// TIA Portal V20 export
// export: Created 2026-10-20T18:54:58.074688Z, ExportSetting None, DisplayName Totally Integrated Automation Portal, DisplayVersion V20 Update 6, DisplayName TIA Portal Openness, DisplayVersion V20 Update 6, DisplayName TIA Portal Version Control Interface, DisplayVersion V20 Update 6, DisplayName SINAMICS Startdrive Advanced, DisplayVersion V20 SP1, DisplayName SINAMICS Startdrive G130, G150, S120, S150, SINAMICS MV, G220, S200, S210, DisplayVersion V20 SP1, DisplayName SINAMICS Startdrive G110M, G120, G120C, G120D, G120P, G115D, DisplayVersion V20 SP1, DisplayName STEP 7 Professional, DisplayVersion V20 Update 6, DisplayName STEP 7 Safety, DisplayVersion V20 Update 2, DisplayName WinCC Basic/Comfort/Advanced, DisplayVersion V20 Update 6, DisplayName WinCC Unified, DisplayVersion V20 Update 6
VAR_GLOBAL   // PLC tag table "IO_ET200_2"
   "C2205 - SENSOR CNV RIGHT (PALLET DETECT 1)" AT %I354.4 : Bool;
   "C2204 - SENSOR CNV RIGHT (PALLET DETECT 1)" AT %I352.4 : Bool;
   "C2206 - SENSOR CNV RIGHT (PALLET DETECT 1)" AT %I356.4 : Bool;
   "C2203 - SENSOR CNV RIGHT (PALLET DETECT 1)" AT %I350.4 : Bool;
   "C2208 - SENSOR CNV RIGHT (PALLET DETECT 1)" AT %I360.4 : Bool;
   "KEY REMOTE/LOCAL L7 - CH2(2)" AT %I1654.5 : Bool;
   "E-STOP L7 - CH2(2)" AT %I1654.4 : Bool;
   "KEY REMOTE/LOCAL L8 - CH1(2)" AT %I1654.3 : Bool;
   "KEY REMOTE/LOCAL L6 - CH1(2)" AT %I1646.3 : Bool;
   "KEY REMOTE/LOCAL L7 - CH1(2)" AT %I1654.1 : Bool;
   "KEY REMOTE/LOCAL L2 - CH2(2)" AT %I1476.7 : Bool;
   "E-STOP L3 - CH1(2)" AT %I1638.0 : Bool;
   "KEY REMOTE/LOCAL L3 - CH1(2)" AT %I1638.1 : Bool;
   "E-STOP L4 - CH1(2)" AT %I1638.2 : Bool;
   "KEY REMOTE/LOCAL L4 - CH1(2)" AT %I1638.3 : Bool;
   "E-STOP L3 - CH2(2)" AT %I1638.4 : Bool;
   "KEY REMOTE/LOCAL L3 - CH2(2)" AT %I1638.5 : Bool;
   "E-STOP L4 - CH2(2)" AT %I1638.6 : Bool;
   "KEY REMOTE/LOCAL L4 - CH2(2)" AT %I1638.7 : Bool;
   "E-STOP L5 - CH1(2)" AT %I1646.0 : Bool;
   "KEY REMOTE/LOCAL L5 - CH1(2)" AT %I1646.1 : Bool;
   "E-STOP L6 - CH1(2)" AT %I1646.2 : Bool;
   "E-STOP L5 - CH2(2)" AT %I1646.4 : Bool;
   "KEY REMOTE/LOCAL L5 - CH2(2)" AT %I1646.5 : Bool;
   "E-STOP L6 - CH2(2)" AT %I1646.6 : Bool;
   "KEY REMOTE/LOCAL L6 - CH2(2)" AT %I1646.7 : Bool;
   "E-STOP L7 - CH1(2)" AT %I1654.0 : Bool;
   "E-STOP L8 - CH1(2)" AT %I1654.2 : Bool;
   "E-STOP L2 - CH2(2)" AT %I1476.6 : Bool;
   "KEY REMOTE/LOCAL L2 - CH1(2)" AT %I1476.3 : Bool;
   "E-STOP L2 - CH1(2)" AT %I1476.2 : Bool;
   "E-STOP L8 - CH2(2)" AT %I1654.6 : Bool;
   "KEY REMOTE/LOCAL L8 - CH2(2)" AT %I1654.7 : Bool;
   "C2102 - SENSOR SAFETY PIN1 DOWN" AT %I175.3 : Bool;
   "C2202 - SENSOR CNV LEFT (PALLET DETECT 2)" AT %I270.0 : Bool;
   "CVTD2 SENSOR CONVEYOR CENTER" AT %I1275.5 : Bool;
   "C2206 - SHUTTLE IN POSITION 2" AT %I357.6 : Bool;
   "C2205 - SENSOR SAFETY PIN1 DOWN" AT %I355.3 : Bool;
   "C2105 - SENSOR CNV LEFT (PALLET DETECT 1)" AT %I194.4 : Bool;
   "C2201 - SENSOR CNV RIGHT" AT %I202.5 : Bool;
   "C2203 - SENSOR CNV LEFT (PALLET DETECT 2)" AT %I351.0 : Bool;
   "C2106 - SENSOR CNV LEFT (PALLET DETECT 2)" AT %I197.1 : Bool;
   "C2107 - SENSOR CNV LEFT" AT %I198.5 : Bool;
   "C2104 - SENSOR CNV LEFT (PALLET DETECT 1)" AT %I178.6 : Bool;
   "C2106 - SENSOR SAFETY PIN1 UP" AT %I197.2 : Bool;
   "C2105 - SENSOR CNV RIGHT (PALLET DETECT 2)" AT %I195.0 : Bool;
   "C2102 - SENSOR CNV LEFT (PALLET DETECT 1)" AT %I174.4 : Bool;
   "C2105 - SENSOR CNV LEFT (PALLET DETECT 2)" AT %I195.1 : Bool;
   "C2106 - SENSOR CNV RIGHT" AT %I197.4 : Bool;
   "VTD2 LEVEL DETECT 1" AT %I1276.7 : Bool;
   "C2206 - SENSOR CNV RIGHT" AT %I356.5 : Bool;
   "C2203 - SENSOR SAFETY PIN1 DOWN" AT %I351.3 : Bool;
   "C2207 - SENSOR SAFETY PIN1 UP" AT %I359.2 : Bool;
   "C2202 - SENSOR CNV LEFT" AT %I270.4 : Bool;
   "C2106 - SENSOR CNV RIGHT (PALLET DETECT 2)" AT %I197.0 : Bool;
   "C2207 - SENSOR CNV RIGHT (PALLET DETECT 2)" AT %I359.1 : Bool;
   "C2203 - SENSOR CNV RIGHT" AT %I350.5 : Bool;
   "C2201 - SHUTTLE IN POSITION 1" AT %I203.7 : Bool;
   "C2105 - SENSOR CNV RIGHT" AT %I195.4 : Bool;
   "C2102 - SHUTTLE IN POSITION 2" AT %I175.6 : Bool;
   "C2206 - SENSOR CNV LEFT" AT %I357.4 : Bool;
   "C2103 - SENSOR CNV LEFT" AT %I177.3 : Bool;
   "C2107 - SENSOR CNV LEFT (PALLET DETECT 2)" AT %I199.1 : Bool;
   "C2204 - SENSOR CNV RIGHT (PALLET DETECT 2)" AT %I353.1 : Bool;
   "C2108 - SHUTTLE IN POSITION 2" AT %I201.6 : Bool;
   "CVTD2 SENSOR CONVEYOR RIGHT" AT %I1275.3 : Bool;
   "C2104 - SENSOR CNV RIGHT (PALLET DETECT 1)" AT %I179.5 : Bool;
   "C2204 - SENSOR CNV LEFT" AT %I353.4 : Bool;
   "C2204 - SENSOR CNV LEFT (PALLET DETECT 2)" AT %I353.0 : Bool;
   "VTD2 ULTIMATE CREEP" AT %I1276.5 : Bool;
   "C2201 - SENSOR CNV RIGHT (PALLET DETECT 2)" AT %I203.1 : Bool;
   "VTD2 DOCKING PINS RETRACTED 1" AT %I1276.2 : Bool;
   "C2201 - SENSOR CNV LEFT (PALLET DETECT 1)" AT %I203.5 : Bool;
   "C2105 - SENSOR SAFETY PIN1 UP" AT %I195.2 : Bool;
   "C2108 - SENSOR CNV LEFT (PALLET DETECT 1)" AT %I200.4 : Bool;
   "C2202 - SENSOR CNV RIGHT (PALLET DETECT 2)" AT %I270.1 : Bool;
   "C2208 - SENSOR CNV LEFT" AT %I361.4 : Bool;
   "C2104 - SENSOR CNV LEFT" AT %I178.7 : Bool;
   "C2107 - SHUTTLE IN POSITION 1" AT %I199.2 : Bool;
   "C2106 - SENSOR SAFETY PIN1 DOWN" AT %I197.3 : Bool;
   "C2206 - SHUTTLE IN POSITION 1" AT %I357.7 : Bool;
   "C2206 - SENSOR CNV RIGHT (PALLET DETECT 2)" AT %I357.1 : Bool;
   "C2107 - SENSOR SAFETY PIN1 UP" AT %I199.7 : Bool;
   "C2206 - SENSOR SAFETY PIN1 UP" AT %I357.2 : Bool;
   "C2106 - SENSOR CNV LEFT" AT %I196.5 : Bool;
   "C2103 - SENSOR CNV LEFT (PALLET DETECT 1)" AT %I177.2 : Bool;
   "C2201 - SHUTTLE IN POSITION 2" AT %I203.6 : Bool;
   "C2106 - SHUTTLE IN POSITION 1" AT %I197.7 : Bool;
   "C2103 - SENSOR CNV RIGHT (PALLET DETECT 1)" AT %I177.5 : Bool;
   "VTD2 DOCKING PINS EXTENDED 1" AT %I1276.0 : Bool;
   "C2101 - SHUTTLE IN POSITION 2" AT %I172.6 : Bool;
   "C2101 - SENSOR CNV LEFT (PALLET DETECT 2)" AT %I172.3 : Bool;
   "C2207 - SENSOR CNV RIGHT" AT %I358.5 : Bool;
   "C2207 - SHUTTLE IN POSITION 2" AT %I359.6 : Bool;
   "C2202 - SENSOR CNV LEFT (PALLET DETECT 1)" AT %I270.5 : Bool;
   "C2102 - SENSOR SAFETY PIN1 UP" AT %I175.2 : Bool;
   "C2101 - SENSOR CNV RIGHT (PALLET DETECT 2)" AT %I172.2 : Bool;
   "C2204 - SENSOR CNV RIGHT" AT %I352.5 : Bool;
   "C2207 - SHUTTLE IN POSITION 1" AT %I359.7 : Bool;
   "C2204 - SHUTTLE IN POSITION 2" AT %I353.6 : Bool;
   "C2203 - SHUTTLE IN POSITION 1" AT %I351.7 : Bool;
   "C2205 - SENSOR CNV RIGHT" AT %I354.5 : Bool;
   "C2202 - SENSOR CNV RIGHT (PALLET DETECT 1)" AT %I269.4 : Bool;
   "C2208 - SENSOR SAFETY PIN1 UP" AT %I361.2 : Bool;
   "C2204 - SENSOR SAFETY PIN1 UP" AT %I353.2 : Bool;
   "C2104 - SHUTTLE IN POSITION 1" AT %I179.7 : Bool;
   "C2101 - SENSOR CNV RIGHT (PALLET DETECT 1)" AT %I172.1 : Bool;
   "C2103 - SENSOR CNV RIGHT" AT %I177.4 : Bool;
   "C2207 - SENSOR CNV RIGHT (PALLET DETECT 1)" AT %I358.4 : Bool;
   "C2204 - SENSOR SAFETY PIN1 DOWN" AT %I353.3 : Bool;
   "C2107 - SENSOR CNV RIGHT (PALLET DETECT 2)" AT %I199.0 : Bool;
   "C2106 - SHUTTLE IN POSITION 2" AT %I197.6 : Bool;
   "C2208 - SHUTTLE IN POSITION 1" AT %I361.7 : Bool;
   "C2208 - SENSOR CNV LEFT (PALLET DETECT 2)" AT %I361.0 : Bool;
   "C2208 - SENSOR CNV RIGHT (PALLET DETECT 2)" AT %I361.1 : Bool;
   "C2104 - SENSOR SAFETY PIN1 UP" AT %I179.2 : Bool;
   "C2202 - SHUTTLE IN POSITION 1" AT %I270.7 : Bool;
   "C2202 - SENSOR CNV RIGHT" AT %I269.5 : Bool;
   "C2205 - SENSOR SAFETY PIN1 UP" AT %I355.2 : Bool;
   "C2201 - SENSOR CNV RIGHT (PALLET DETECT 1)" AT %I202.4 : Bool;
   "C2205 - SHUTTLE IN POSITION 2" AT %I355.6 : Bool;
   "C2202 - SHUTTLE IN POSITION 2" AT %I270.6 : Bool;
   "C2201 - SENSOR CNV LEFT" AT %I203.4 : Bool;
   "C2207 - SENSOR SAFETY PIN1 DOWN" AT %I359.3 : Bool;
   "C2207 - SENSOR CNV LEFT" AT %I359.4 : Bool;
   "C2101 - SENSOR CNV RIGHT" AT %I172.0 : Bool;
   "C2102 - SENSOR CNV LEFT (PALLET DETECT 2)" AT %I175.1 : Bool;
   "VTD2 ULTIMATE SLOWDOWN" AT %I1276.4 : Bool;
   "C2104 - SENSOR CNV LEFT (PALLET DETECT 2)" AT %I179.1 : Bool;
   "C2106 - SENSOR CNV LEFT (PALLET DETECT 1)" AT %I196.4 : Bool;
   "C2107 - SHUTTLE IN POSITION 2" AT %I199.6 : Bool;
   "C2203 - SENSOR SAFETY PIN1 UP" AT %I351.2 : Bool;
   "C2207 - SENSOR CNV LEFT (PALLET DETECT 2)" AT %I359.0 : Bool;
   "VTD2 DOCKING PINS EXTENDED 2" AT %I1276.1 : Bool;
   "C2201 - SENSOR CNV LEFT (PALLET DETECT 2)" AT %I203.0 : Bool;
   "C2108 - SHUTTLE IN POSITION 1" AT %I201.7 : Bool;
   "C2101 - SENSOR CNV LEFT" AT %I172.5 : Bool;
   "C2107 - SENSOR CNV RIGHT (PALLET DETECT 1)" AT %I199.5 : Bool;
   "C2203 - SHUTTLE IN POSITION 2" AT %I351.6 : Bool;
   "C2107 - SENSOR CNV LEFT (PALLET DETECT 1)" AT %I198.4 : Bool;
   "C2208 - SHUTTLE IN POSITION 2" AT %I361.6 : Bool;
   "C2205 - SENSOR CNV LEFT" AT %I355.4 : Bool;
   "C2203 - SENSOR CNV LEFT" AT %I351.4 : Bool;
   "C2105 - SENSOR CNV RIGHT (PALLET DETECT 1)" AT %I195.5 : Bool;
   "C2108 - SENSOR CNV RIGHT" AT %I201.4 : Bool;
   "C2108 - SENSOR CNV RIGHT (PALLET DETECT 2)" AT %I201.0 : Bool;
   "C2208 - SENSOR SAFETY PIN1 DOWN" AT %I361.3 : Bool;
   "C2104 - SHUTTLE IN POSITION 2" AT %I179.6 : Bool;
   "C2101 - SENSOR CNV LEFT (PALLET DETECT 1)" AT %I172.4 : Bool;
   "C2102 - SENSOR CNV RIGHT (PALLET DETECT 2)" AT %I175.0 : Bool;
   "C2105 - SHUTTLE IN POSITION 2" AT %I195.6 : Bool;
   "C2103 - SENSOR CNV LEFT (PALLET DETECT 2)" AT %I177.1 : Bool;
   "C2203 - SENSOR CNV LEFT (PALLET DETECT 1)" AT %I351.5 : Bool;
   "C2103 - SHUTTLE IN POSITION 2" AT %I177.6 : Bool;
   "C2106 - SENSOR CNV RIGHT (PALLET DETECT 1)" AT %I197.5 : Bool;
   "CVTD2 SENSOR CONVEYOR LEFT (PALLET DETECT 1)" AT %I1275.2 : Bool;
   "C2105 - SHUTTLE IN POSITION 1" AT %I195.7 : Bool;
   "C2102 - SENSOR CNV LEFT" AT %I174.5 : Bool;
   "VTD2 DOCKING PINS RETRACTED 2" AT %I1276.3 : Bool;
   "VTD2 LEVEL DETECT 2" AT %I1276.6 : Bool;
   "C2203 - SENSOR CNV RIGHT (PALLET DETECT 2)" AT %I351.1 : Bool;
   "C2103 - SENSOR CNV RIGHT (PALLET DETECT 2)" AT %I177.0 : Bool;
   "C2206 - SENSOR SAFETY PIN1 DOWN" AT %I357.3 : Bool;
   "C2206 - SENSOR CNV LEFT (PALLET DETECT 1)" AT %I357.5 : Bool;
   "C2205 - SENSOR CNV LEFT (PALLET DETECT 1)" AT %I355.5 : Bool;
   "C2205 - SENSOR CNV RIGHT (PALLET DETECT 2)" AT %I355.1 : Bool;
   "CVTD2 SENSOR CONVEYOR LEFT" AT %I1275.1 : Bool;
   "C2102 - SENSOR CNV RIGHT" AT %I175.4 : Bool;
   "C2204 - SENSOR CNV LEFT (PALLET DETECT 1)" AT %I353.5 : Bool;
   "C2208 - SENSOR CNV RIGHT" AT %I360.5 : Bool;
   "C2205 - SENSOR CNV LEFT (PALLET DETECT 2)" AT %I355.0 : Bool;
   "C2107 - SENSOR SAFETY PIN1 DOWN" AT %I199.3 : Bool;
   "C2107 - SENSOR CNV RIGHT" AT %I199.4 : Bool;
   "C2101 - SHUTTLE IN POSITION 1" AT %I172.7 : Bool;
   "C2208 - SENSOR CNV LEFT (PALLET DETECT 1)" AT %I361.5 : Bool;
   "C2205 - SHUTTLE IN POSITION 1" AT %I355.7 : Bool;
   "C2104 - SENSOR CNV RIGHT" AT %I179.4 : Bool;
   "C2202 - SENSOR SAFETY PIN1 UP" AT %I270.2 : Bool;
   "C2103 - SHUTTLE IN POSITION 1" AT %I177.7 : Bool;
   "C2204 - SHUTTLE IN POSITION 1" AT %I353.7 : Bool;
   "C2104 - SENSOR SAFETY PIN1 DOWN" AT %I179.3 : Bool;
   "C2202 - SENSOR SAFETY PIN1 DOWN" AT %I270.3 : Bool;
   "C2104 - SENSOR CNV RIGHT (PALLET DETECT 2)" AT %I179.0 : Bool;
   "C2206 - SENSOR CNV LEFT (PALLET DETECT 2)" AT %I357.0 : Bool;
   "C2102 - SENSOR CNV RIGHT (PALLET DETECT 1)" AT %I175.5 : Bool;
   "C2105 - SENSOR CNV LEFT" AT %I194.5 : Bool;
   "C2102 - SHUTTLE IN POSITION 1" AT %I175.7 : Bool;
   "C2105 - SENSOR SAFETY PIN1 DOWN" AT %I195.3 : Bool;
   "C2207 - SENSOR CNV LEFT (PALLET DETECT 1)" AT %I359.5 : Bool;
   "C2108 - SENSOR CNV RIGHT (PALLET DETECT 1)" AT %I201.5 : Bool;
   "CVTD2 SENSOR CONVEYOR RIGHT (PALLET DETECT 1)" AT %I1275.4 : Bool;
   "C2103 - SENSOR SAFETY PIN1 DOWN" AT %I176.5 : Bool;
   "C2103 - SENSOR SAFETY PIN1 UP" AT %I176.4 : Bool;
   "C2108 - SENSOR SAFETY PIN1 UP" AT %I201.2 : Bool;
   "C2108 - SENSOR SAFETY PIN1 DOWN" AT %I201.3 : Bool;
   "C2108 - SENSOR CNV LEFT" AT %I200.5 : Bool;
   "C2108 - SENSOR CNV LEFT (PALLET DETECT 2)" AT %I201.1 : Bool;
   "KEY REMOTE/LOCAL L1 - CH1(2)" AT %I1476.0 : Bool;
   "E-STOP L1 - CH1(2)" AT %I1476.1 : Bool;
   "KEY REMOTE/LOCAL L1 - CH2(2)" AT %I1476.4 : Bool;
   "E-STOP L1 - CH2(2)" AT %I1476.5 : Bool;
   "CVTD2 OVERHANG LEFT" AT %I1275.6 : Bool;
   "CVTD2 OVERHANG RIGHT" AT %I1275.7 : Bool;
END_VAR
